Fanuc KAREL source: kb00087.KL

-- PROVISIONAL review KL for V940-1; original PC SHA256 e4421528e13d1873fe3c32613a342955e9dfd995317de2fe0f01f0d5e7303e38
-- Incomplete behavior may be omitted. Consult companion uncertainty JSON. Do not deploy.
PROGRAM KB00087
%NOLOCKGROUP
BEGIN
  -- V9_ZERO_TABLE_METADATA_HINT layout=0002_ascii; no indexed target words; source/name/runtime held
  -- UNRESOLVED_PC offsets 5-12; opcodes 9D,23
  -- UNRESOLVED_PC offsets 17-24; opcodes 9D,23
  -- UNRESOLVED_PC offsets 29-59; opcodes 27,22,22,27,9D,31,7E,4A
  -- UNRESOLVED_PC offsets 64-68; opcodes 7F
END KB00087
